{attribute 'qualified_only'}
{attribute 'strict'}
{attribute 'to_string'}
TYPE E_LogRecordQueueFailureReason :
(
	NA := 0,  // No failure occurred.
	RECORD_POINTER_NULL,  // The supplied log-record pointer is null.
	DESTINATION_ALREADY_ASSIGNED,  // The pop destination pointer is already assigned.
	QUEUE_EMPTY,  // The queue contains no record to pop.
	MAX_SIZE_ENFORCEMENT_FAILURE := 5,  // The bounded eviction loop could not restore the configured maximum size.
	DESTINATION_NOT_EMPTY,  // The transfer destination already owns records.
	DESTINATION_CAPACITY_TOO_SMALL,  // The transfer destination cannot hold every source record.
	SELF_TRANSFER_NOT_ALLOWED,  // A queue cannot transfer ownership to itself.
	MEMORY_ALLOCATION_FAILURE  // Dynamic node allocation failed.
) UDINT;
END_TYPE

(* stored: Version 1.1.0.1
   EnumerationTextList E_LogRecordQueueFailureReason: Id {889b75ee-4565-4114-a653-39ae2d0d3f52} *)
